Staubli VAL3: Lab2A_L2.dtx


